(*
SPDX-FileCopyrightText: © 2026 Oleksandr Tiutyk <trofimich@gmail.com>
SPDX-License-Identifier: MIT
License: https://opensource.org/license/mit
*)

(*
Catches a framework exception and copies its diagnostic into an ERROR snapshot.

Write _RunRequested once. The sample deliberately raises a standard exception, captures it in the same scan,
and keeps the copied diagnostic after transient exception cleanup. Watch _Error.TopMessage.
Map this program to one dedicated cyclic task. The program performs cleanup for that task.
*)

{attribute 'no_explicit_call' := 'do not call this function block directly'}
PROGRAM ExceptionSnapshotExample
VAR
	{attribute 'hide'}
	_ClassName : STRING := __POUNAME();
	_RunRequested : BOOL;
	_Error : TOF_Core.ERROR;
END_VAR

TOF_Core.System.Execute();

IF _RunRequested THEN
	_RunRequested := FALSE;
	captureExampleError();
END_IF

TOF_Core.DynamicMemoryManager.RaiseIfAllocationFailed();
TOF_Core.DynamicMemoryManager.CleanupMemory();

// Copies the demonstration failure before the task cleans up the exception.
METHOD PRIVATE captureExampleError
VAR
	exceptionCode : __SYSTEM.ExceptionCode;
	caught : TOF_Core.IException;
END_VAR
_Error.Clear();

__TRY
	TOF_Core.Exceptions.ThrowStandard(
		sourceNamespaceName := NamespaceName,
		sourceClassName := ClassName,
		sourcePOUName := __POUNAME(),
		sourcePosition := __POSITION(),
		message := "Example operation failed"
	);
__CATCH(exceptionCode)
	caught := TOF_Core.ExceptionManager.GetLastException(
		exceptionCode := exceptionCode,
		catchPointNamespaceName := NamespaceName,
		catchPointPOUName := __POUNAME(),
		catchPointPosition := __POSITION()
	);
	caught.ToError(targetError := _Error, severity := TOF_Core.ERROR_SEVERITY.ERROR);
__ENDTRY
END_METHOD

// Borrows the initialized program name. Treat it as read-only.
{attribute 'monitoring' := 'call'}
PROPERTY ClassName : REFERENCE TO STRING
GET
ClassName REF= _ClassName;
END_GET
END_PROPERTY

// Borrows the initialized namespace name. Treat it as read-only.
{attribute 'monitoring' := 'call'}
PROPERTY NamespaceName : REFERENCE TO STRING
GET
NamespaceName REF= CurrentNamespace.Name;
END_GET
END_PROPERTY

END_PROGRAM

(* stored: Version 1.1.0.1
   POU ExceptionSnapshotExample: Id {6f4a565e-cfa2-433b-832e-adb6cabe01fc}, SpecialFunc None
   Method captureExampleError: Id {4294fd11-78cb-4baa-9406-6a6a107d1559}
   Property ClassName: Id {afed3e86-f5e7-41a5-925e-7ec67182d41e}
   Get Get: Id {e49c0505-45bb-4fdd-aad6-9f2b8fc427ac}
   Property NamespaceName: Id {337e7e3f-18e7-4454-aaff-7329285bb44e}
   Get Get: Id {fba8a079-ae65-424d-894c-451cd5143b84} *)
